TYPE ST_FeedConfig :
STRUCT
    sId           : STRING(20);     // short id used in the payloads: F1, F2
    sName         : STRING(40);
    fMaxAmps      : LREAL := 32.0;  // A per leg
    fWireLengthFt : LREAL := 0.0;   // one-way length of the infeed cable: meter to the point where the boxes branch off
    nWireAwg      : INT := 10;      // AWG of one conductor, copper
END_STRUCT
END_TYPE

(* stored: Version 1.1.0.1
   DUT ST_FeedConfig: Id {18adeafb-2171-4642-893d-1330bbb7dac6} *)
